(* Logix 5000 project; controller R400_500_XLS vendor 1 type 14 code 216 rev 31.11; software revision 31.01; part 12 of 32 *)
(* tags used below, declared in another part *)
   Chem_Pump : UDT_CHEM_PUMP[4];   // Chemical Pump flow rate
   CHEMICAL_COND_MAX_TIME : DINT;   // Timeout for the conductivity based chemical injection
   CHEMICAL_PUMP_OFF_TIME : DINT[4];
   CHEMICAL_PUMP_ON_TIME : DINT[4];
   FC87_CalibChemPmp : SINT;   // Calibration chemical pumps activation bits
   FC87_CalibChemPmpMsg : SINT;   // Chemical pump calibration step message
   FC87_ChemCalibRemainTime : DINT;
   FC87_ChemPumpIndex : SINT;   // Index of the selected chemical pump to calibrate
   FC87_LastValue : SINT;
   FC87_ONS : DINT;
   M : DINT[5];   // Memory Bits
   ONS_SPV17 : SINT;
   SET_POINT_FRACTION : REAL[4];
   Supervisor : DINT;
   Tmr : TIMER[107];
   ChemicalName : STRING[9];   // Used by HMI
   ChemPumpSelector : UDT_SELECTOR[2];   // Chemical pump calibration selector
   Current_Screen : DINT;
   DateTime : DINT[7];
   DateTimeNew : DINT[7];
   NumInput : UDT_NUMERIC_INPUT[65];   // Numeric input
   NumInputReal : UDT_NUMERIC_INPUT_REAL[17];
   RemoteDayOfMonth : DINT;   // HMI Date Day
   RemoteHour : DINT;   // HMI Time Hour
   RemoteMinute : DINT;   // HMI Time Minute
   RemoteMonth : DINT;   // HMI Date Month
   RemoteSecond : DINT;   // HMI Time Second
   RemoteSetDateTime : BOOL;   // HMI Set Date and Time
   RemoteYear : DINT;   // HMI Date Year
   Screen_Ctrl : DINT;   // PLC Screen Request
   SelChemi_Remote : SINT;
   SelChemical_Ind : SINT;
   SelChemical_Value : SINT;
   Selector : UDT_SELECTOR[25];   // Piloted list selector
   StringInput : UDT_STRING_INPUT[6];
   Tpb : DINT[11];
   TpbImage : DINT[11];
   Unit : Hrdwre;   // Unit Configuration
(* MainProgram, continued *)

ROUTINE SPV_12_CHEM_PUMP_CALIBRATION   (* ladder *)
// Calculate chemical pumps flow rate
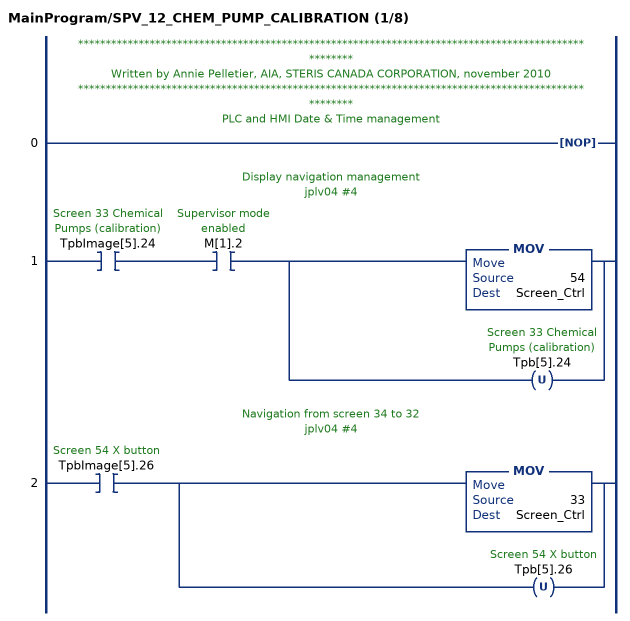
   // ****************************************************************************************************
   // Written by Annie Pelletier, AIA, STERIS CANADA CORPORATION, november 2010
   // ****************************************************************************************************
   // PLC and HMI Date & Time management
   0: NOP();
   // Display navigation management
   // jplv04 #4
   1: XIC(TpbImage[5].24)XIC(M[1].2)[MOV(54,Screen_Ctrl) ,OTU(Tpb[5].24) ];
   // Navigation from screen 34 to 32
   // jplv04 #4
   2: XIC(TpbImage[5].26)[MOV(33,Screen_Ctrl) ,OTU(Tpb[5].26) ];
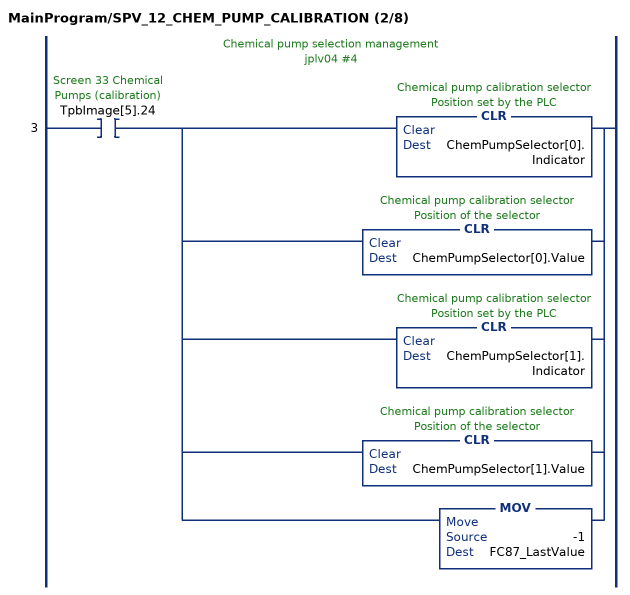
   // Chemical pump selection management
   // jplv04 #4
   3: XIC(TpbImage[5].24)[CLR(ChemPumpSelector[0].Indicator) ,CLR(ChemPumpSelector[0].Value) ,CLR(ChemPumpSelector[1].Indicator) ,CLR(ChemPumpSelector[1].Value) ,MOV(-1,FC87_LastValue) ];
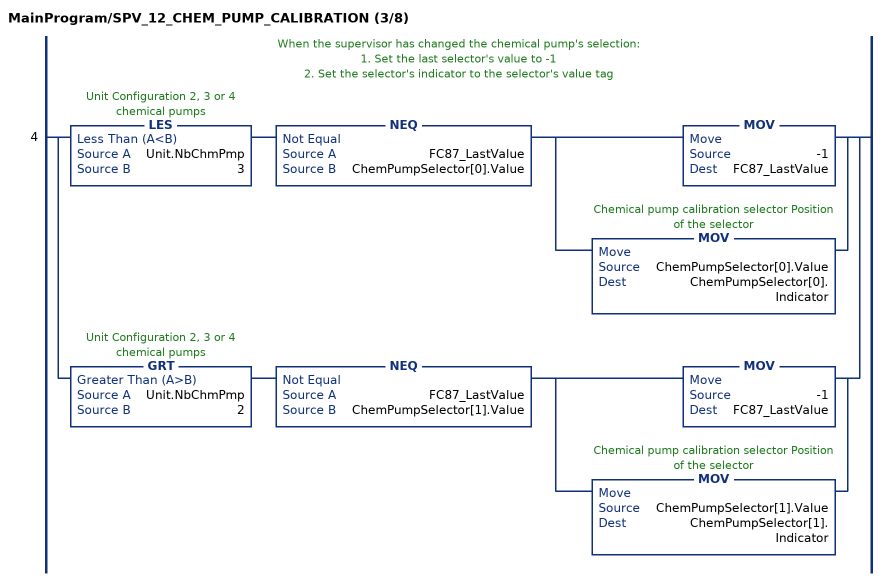
   // When the supervisor has changed the chemical pump's selection:
   // 1. Set the last selector's value to -1
   // 2. Set the selector's indicator to the selector's value tag
   4: [LES(Unit.NbChmPmp,3) NEQ(FC87_LastValue,ChemPumpSelector[0].Value) [MOV(-1,FC87_LastValue) ,MOV(ChemPumpSelector[0].Value,ChemPumpSelector[0].Indicator) ] ,GRT(Unit.NbChmPmp,2) NEQ(FC87_LastValue,ChemPumpSelector[1].Value) [MOV(-1,FC87_LastValue) ,MOV(ChemPumpSelector[1].Value,ChemPumpSelector[1].Indicator) ] ];
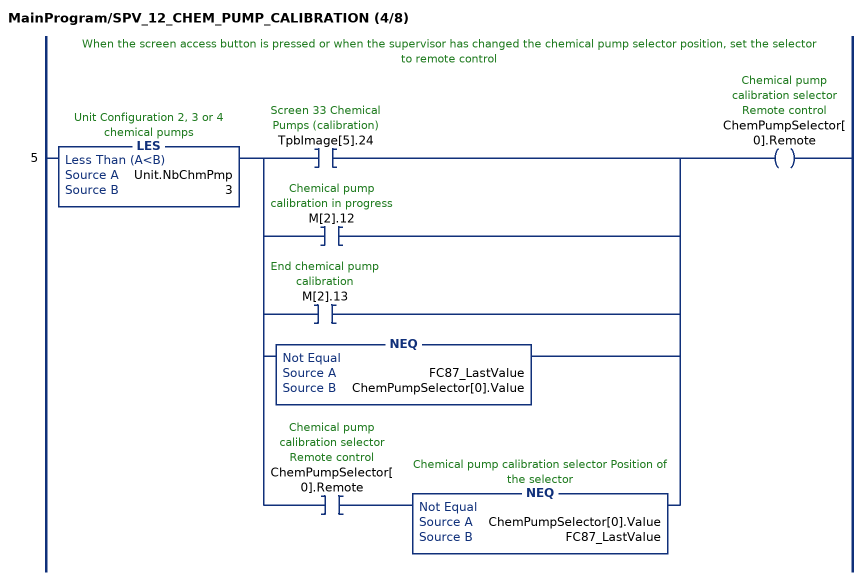
   // When the screen access button is pressed or when the supervisor has changed the chemical pump selector position, set the selector to remote control
   5: LES(Unit.NbChmPmp,3)[XIC(TpbImage[5].24) ,XIC(M[2].12) ,XIC(M[2].13) ,NEQ(FC87_LastValue,ChemPumpSelector[0].Value) ,XIC(ChemPumpSelector[0].Remote) NEQ(ChemPumpSelector[0].Value,FC87_LastValue) ]OTE(ChemPumpSelector[0].Remote);
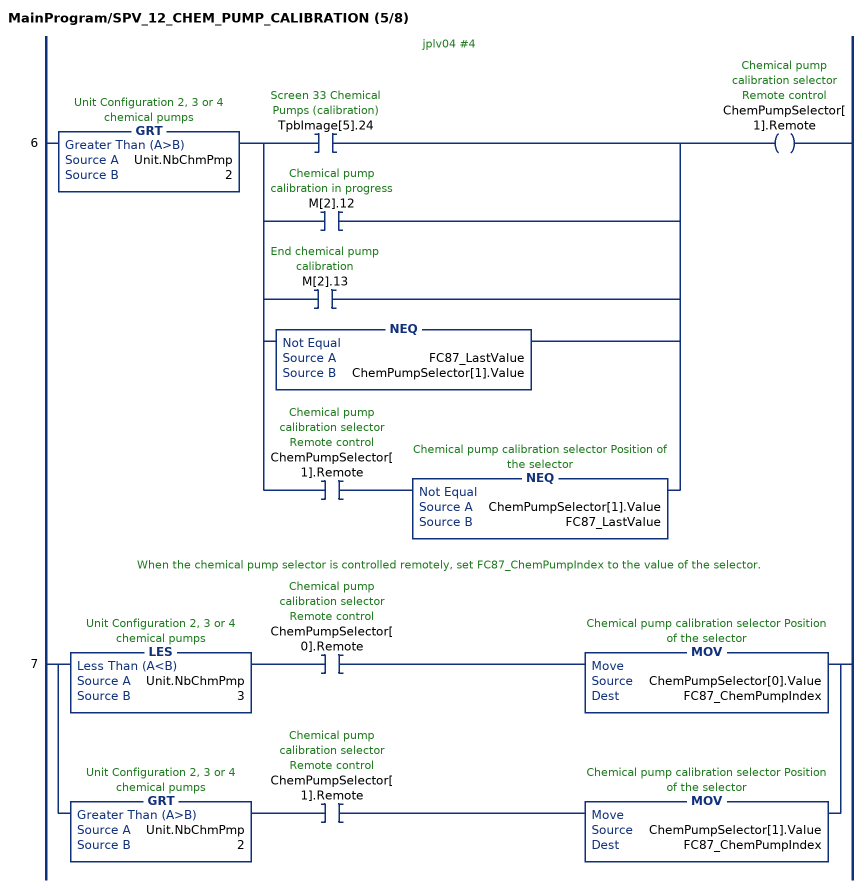
   // jplv04 #4
   6: GRT(Unit.NbChmPmp,2)[XIC(TpbImage[5].24) ,XIC(M[2].12) ,XIC(M[2].13) ,NEQ(FC87_LastValue,ChemPumpSelector[1].Value) ,XIC(ChemPumpSelector[1].Remote) NEQ(ChemPumpSelector[1].Value,FC87_LastValue) ]OTE(ChemPumpSelector[1].Remote);
   // When the chemical pump selector is controlled remotely, set FC87_ChemPumpIndex to the value of the selector.
   7: [LES(Unit.NbChmPmp,3) XIC(ChemPumpSelector[0].Remote) MOV(ChemPumpSelector[0].Value,FC87_ChemPumpIndex) ,GRT(Unit.NbChmPmp,2) XIC(ChemPumpSelector[1].Remote) MOV(ChemPumpSelector[1].Value,FC87_ChemPumpIndex) ];
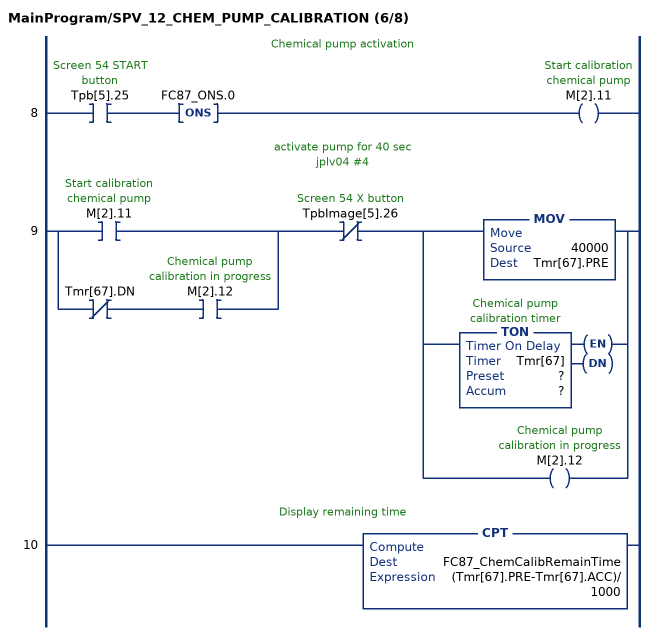
   // Chemical pump activation
   8: XIC(Tpb[5].25)ONS(FC87_ONS.0)OTE(M[2].11);
   // activate pump for 40 sec
   // jplv04 #4
   9: [XIC(M[2].11) ,XIO(Tmr[67].DN) XIC(M[2].12) ]XIO(TpbImage[5].26)[MOV(40000,Tmr[67].PRE) ,TON(Tmr[67],?,?) ,OTE(M[2].12) ];
   // Display remaining time
   10: CPT(FC87_ChemCalibRemainTime,(Tmr[67].PRE-Tmr[67].ACC)/1000);
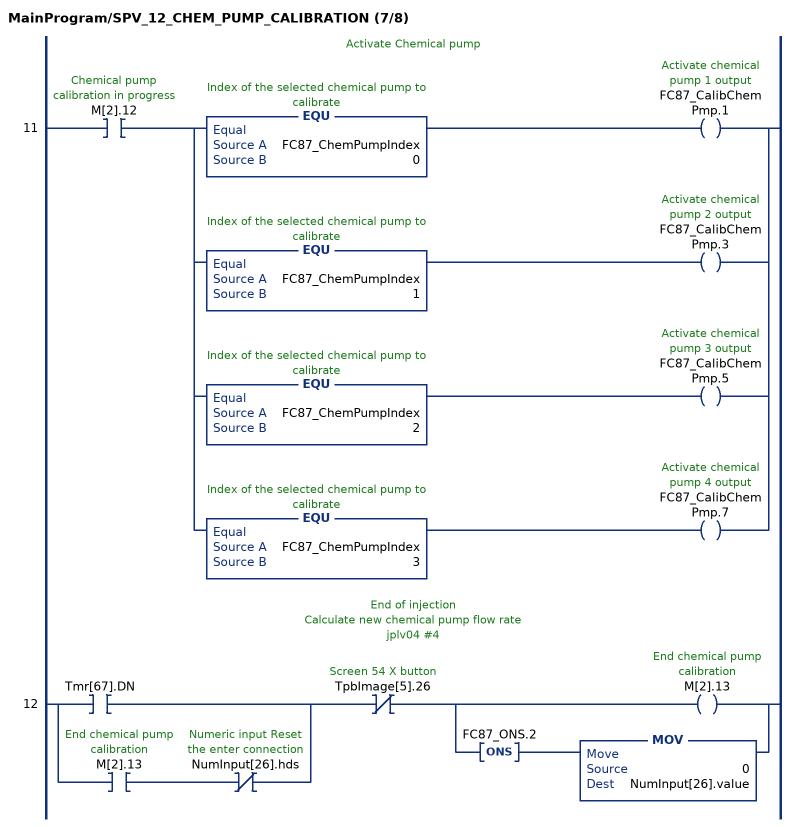
   // Activate Chemical pump
   11: XIC(M[2].12)[EQU(FC87_ChemPumpIndex,0) OTE(FC87_CalibChemPmp.1) ,EQU(FC87_ChemPumpIndex,1) OTE(FC87_CalibChemPmp.3) ,EQU(FC87_ChemPumpIndex,2) OTE(FC87_CalibChemPmp.5) ,EQU(FC87_ChemPumpIndex,3) OTE(FC87_CalibChemPmp.7) ];
   // End of injection
   // Calculate new chemical pump flow rate
   // jplv04 #4
   12: [XIC(Tmr[67].DN) ,XIC(M[2].13) XIO(NumInput[26].hds) ]XIO(TpbImage[5].26)[OTE(M[2].13) ,ONS(FC87_ONS.2) MOV(0,NumInput[26].value) ];
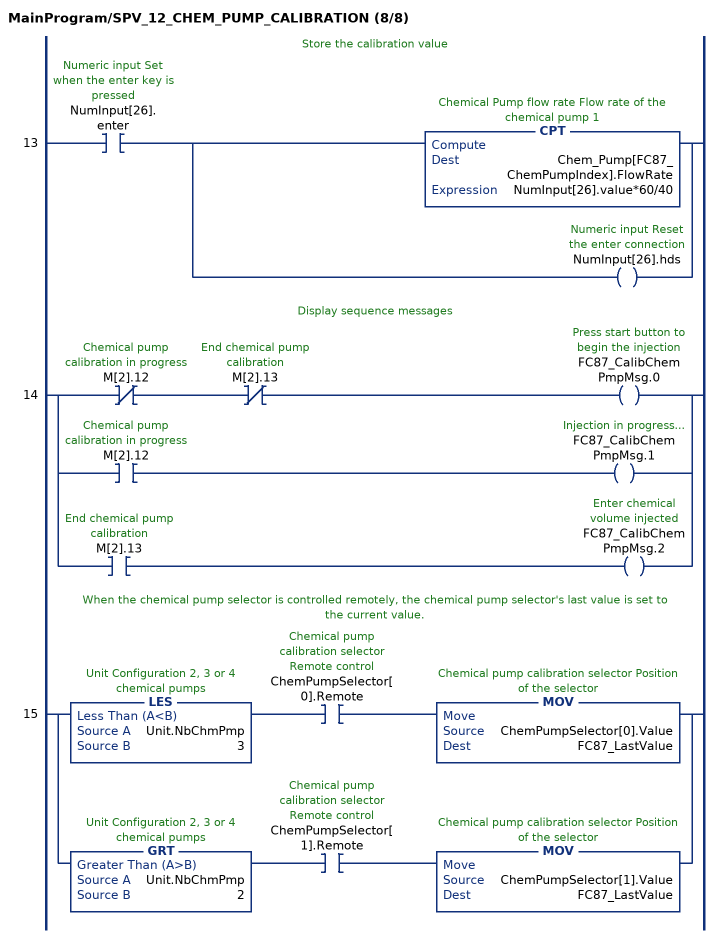
   // Store the calibration value
   13: XIC(NumInput[26].enter)[CPT(Chem_Pump[FC87_ChemPumpIndex].FlowRate,NumInput[26].value*60/40) ,OTE(NumInput[26].hds) ];
   // Display sequence messages
   14: [XIO(M[2].12) XIO(M[2].13) OTE(FC87_CalibChemPmpMsg.0) ,XIC(M[2].12) OTE(FC87_CalibChemPmpMsg.1) ,XIC(M[2].13) OTE(FC87_CalibChemPmpMsg.2) ];
   // When the chemical pump selector is controlled remotely, the chemical pump selector's last value is set to the current value.
   15: [LES(Unit.NbChmPmp,3) XIC(ChemPumpSelector[0].Remote) MOV(ChemPumpSelector[0].Value,FC87_LastValue) ,GRT(Unit.NbChmPmp,2) XIC(ChemPumpSelector[1].Remote) MOV(ChemPumpSelector[1].Value,FC87_LastValue) ];
END_ROUTINE

ROUTINE SPV_16_DATE_TIME   (* ladder *)
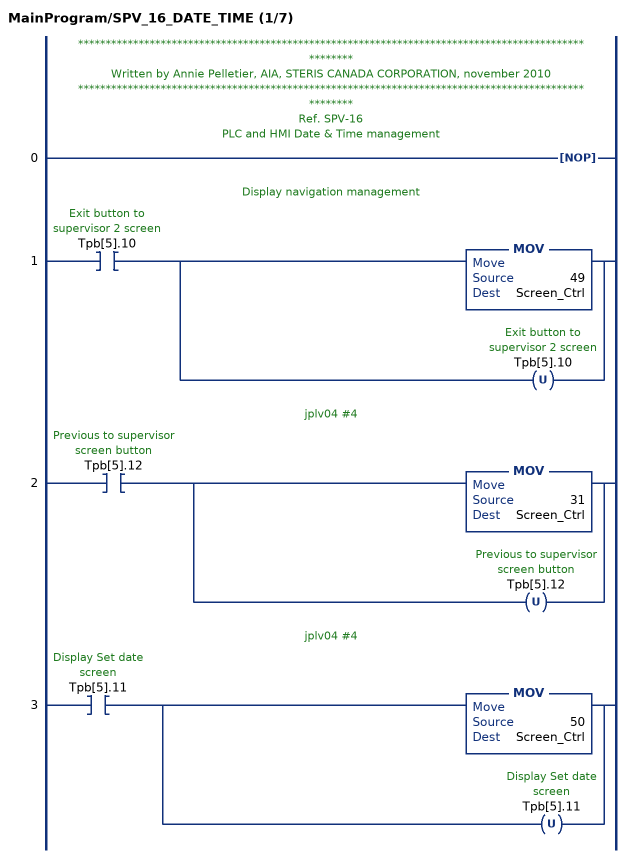
   // ****************************************************************************************************
   // Written by Annie Pelletier, AIA, STERIS CANADA CORPORATION, november 2010
   // ****************************************************************************************************
   // Ref. SPV-16
   // PLC and HMI Date & Time management
   0: NOP();
   // Display navigation management
   1: XIC(Tpb[5].10)[MOV(49,Screen_Ctrl) ,OTU(Tpb[5].10) ];
   // jplv04 #4
   2: XIC(Tpb[5].12)[MOV(31,Screen_Ctrl) ,OTU(Tpb[5].12) ];
   // jplv04 #4
   3: XIC(Tpb[5].11)[MOV(50,Screen_Ctrl) ,OTU(Tpb[5].11) ];
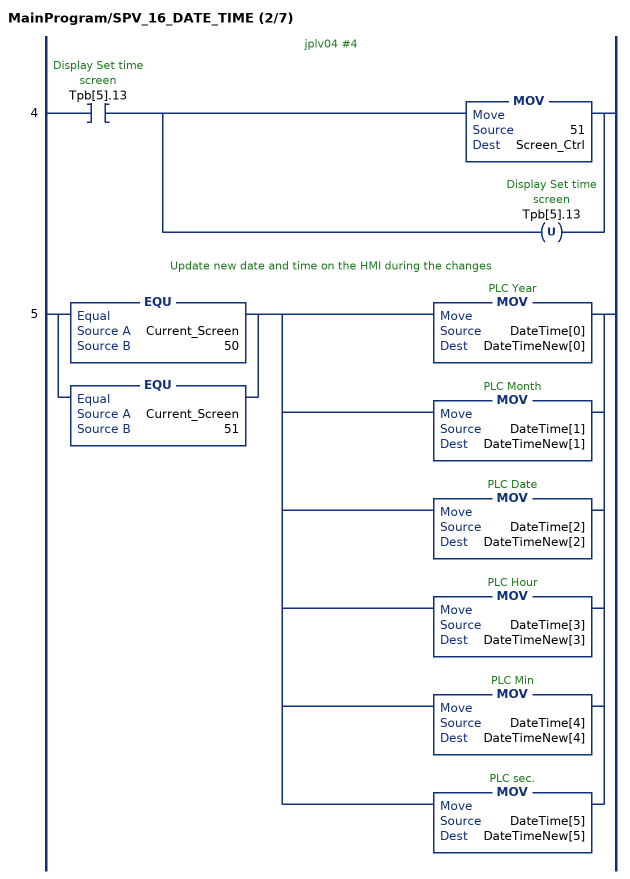
   // jplv04 #4
   4: XIC(Tpb[5].13)[MOV(51,Screen_Ctrl) ,OTU(Tpb[5].13) ];
   // Update new date and time on the HMI during the changes
   5: [EQU(Current_Screen,50) ,EQU(Current_Screen,51) ][MOV(DateTime[0],DateTimeNew[0]) ,MOV(DateTime[1],DateTimeNew[1]) ,MOV(DateTime[2],DateTimeNew[2]) ,MOV(DateTime[3],DateTimeNew[3]) ,MOV(DateTime[4],DateTimeNew[4]) ,MOV(DateTime[5],DateTimeNew[5]) ];
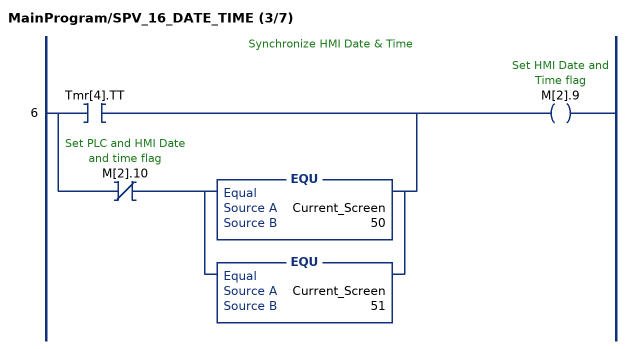
   // Synchronize HMI Date & Time
   6: [XIC(Tmr[4].TT) ,XIO(M[2].10) [EQU(Current_Screen,50) ,EQU(Current_Screen,51) ] ]OTE(M[2].9);
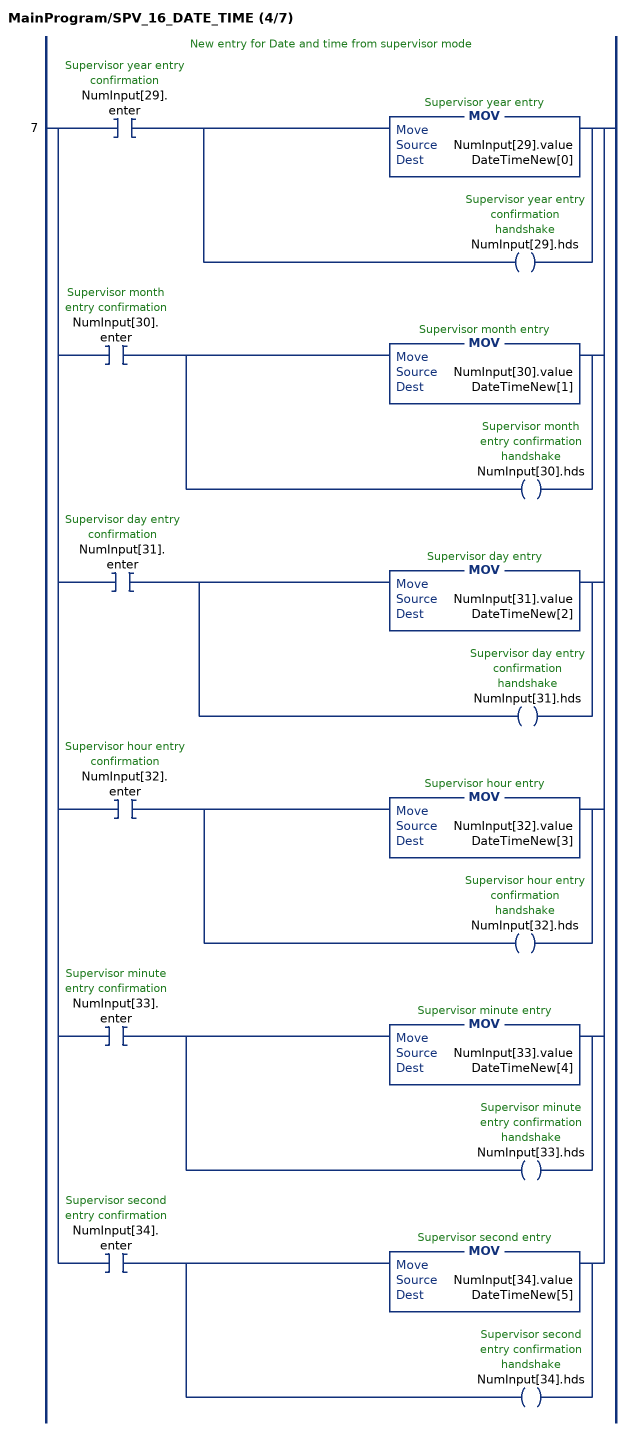
   // New entry for Date and time from supervisor mode
   7: [XIC(NumInput[29].enter) [MOV(NumInput[29].value,DateTimeNew[0]) ,OTE(NumInput[29].hds) ] ,XIC(NumInput[30].enter) [MOV(NumInput[30].value,DateTimeNew[1]) ,OTE(NumInput[30].hds) ] ,XIC(NumInput[31].enter) [MOV(NumInput[31].value,DateTimeNew[2]) ,OTE(NumInput[31].hds) ] ,XIC(NumInput[32].enter) [MOV(NumInput[32].value,DateTimeNew[3]) ,OTE(NumInput[32].hds) ] ,XIC(NumInput[33].enter) [MOV(NumInput[33].value,DateTimeNew[4]) ,OTE(NumInput[33].hds) ] ,XIC(NumInput[34].enter) [MOV(NumInput[34].value,DateTimeNew[5]) ,OTE(NumInput[34].hds) ] ];
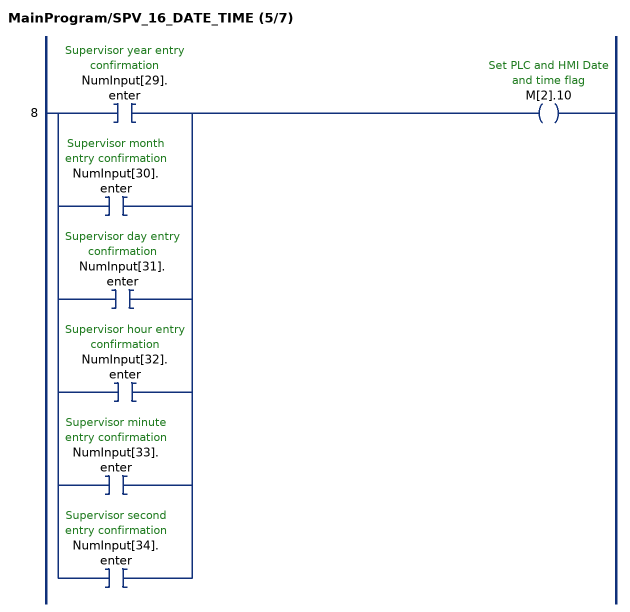
   8: [XIC(NumInput[29].enter) ,XIC(NumInput[30].enter) ,XIC(NumInput[31].enter) ,XIC(NumInput[32].enter) ,XIC(NumInput[33].enter) ,XIC(NumInput[34].enter) ]OTE(M[2].10);
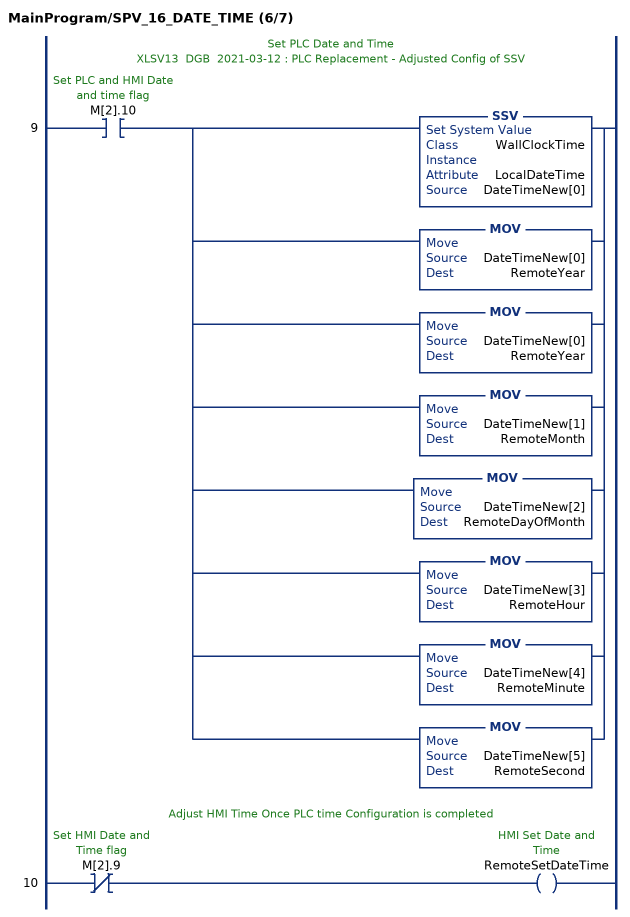
   // Set PLC Date and Time
   // XLSV13  DGB  2021-03-12 : PLC Replacement - Adjusted Config of SSV
   9: XIC(M[2].10)[SSV(WallClockTime,,LocalDateTime,DateTimeNew[0]) ,MOV(DateTimeNew[0],RemoteYear) ,MOV(DateTimeNew[0],RemoteYear) ,MOV(DateTimeNew[1],RemoteMonth) ,MOV(DateTimeNew[2],RemoteDayOfMonth) ,MOV(DateTimeNew[3],RemoteHour) ,MOV(DateTimeNew[4],RemoteMinute) ,MOV(DateTimeNew[5],RemoteSecond) ];
   // Adjust HMI Time Once PLC time Configuration is completed
   10: XIO(M[2].9)OTE(RemoteSetDateTime);
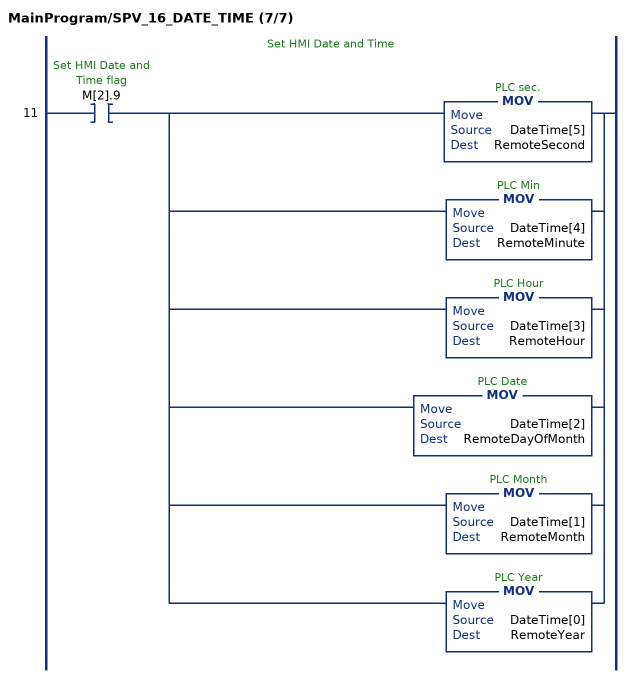
   // Set HMI Date and Time
   11: XIC(M[2].9)[MOV(DateTime[5],RemoteSecond) ,MOV(DateTime[4],RemoteMinute) ,MOV(DateTime[3],RemoteHour) ,MOV(DateTime[2],RemoteDayOfMonth) ,MOV(DateTime[1],RemoteMonth) ,MOV(DateTime[0],RemoteYear) ];
END_ROUTINE

ROUTINE SPV_17_Chemical_Parameters   (* ladder *)
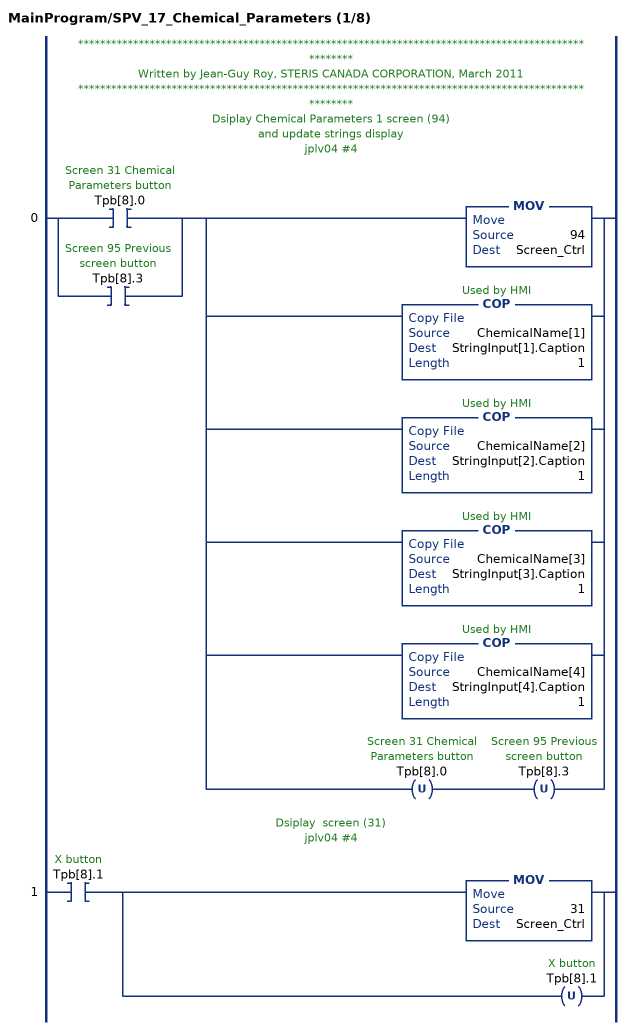
   // ****************************************************************************************************
   // Written by Jean-Guy Roy, STERIS CANADA CORPORATION, March 2011
   // ****************************************************************************************************
   // Dsiplay Chemical Parameters 1 screen (94)
   // and update strings display
   // jplv04 #4
   0: [XIC(Tpb[8].0) ,XIC(Tpb[8].3) ][MOV(94,Screen_Ctrl) ,COP(ChemicalName[1],StringInput[1].Caption,1) ,COP(ChemicalName[2],StringInput[2].Caption,1) ,COP(ChemicalName[3],StringInput[3].Caption,1) ,COP(ChemicalName[4],StringInput[4].Caption,1) ,OTU(Tpb[8].0) OTU(Tpb[8].3) ];
   // Dsiplay  screen (31)
   // jplv04 #4
   1: XIC(Tpb[8].1)[MOV(31,Screen_Ctrl) ,OTU(Tpb[8].1) ];
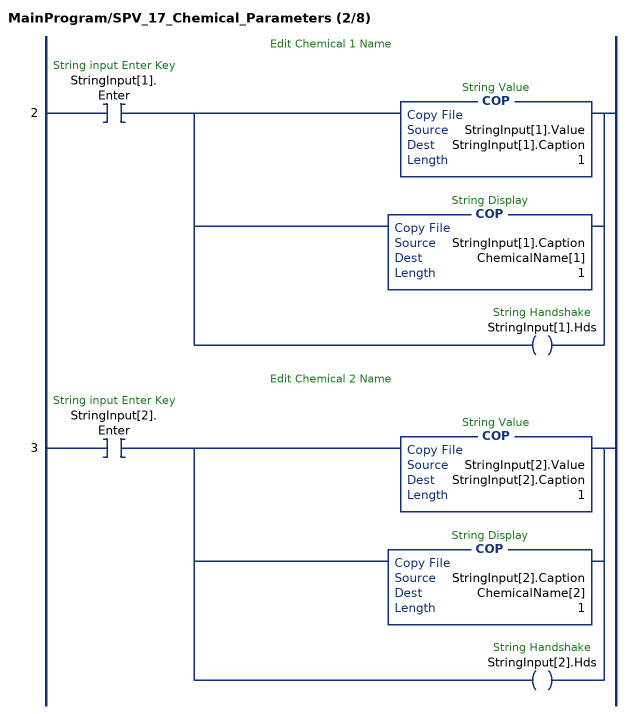
   // Edit Chemical 1 Name
   2: XIC(StringInput[1].Enter)[COP(StringInput[1].Value,StringInput[1].Caption,1) ,COP(StringInput[1].Caption,ChemicalName[1],1) ,OTE(StringInput[1].Hds) ];
   // Edit Chemical 2 Name
   3: XIC(StringInput[2].Enter)[COP(StringInput[2].Value,StringInput[2].Caption,1) ,COP(StringInput[2].Caption,ChemicalName[2],1) ,OTE(StringInput[2].Hds) ];
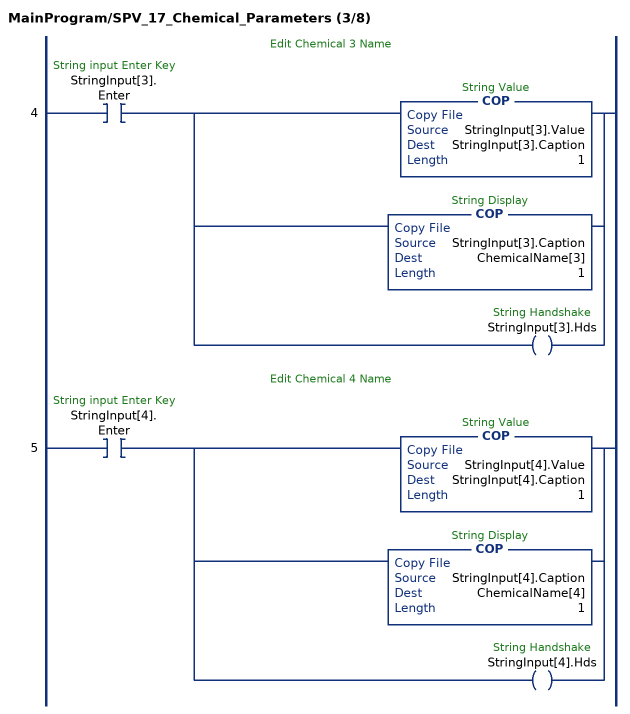
   // Edit Chemical 3 Name
   4: XIC(StringInput[3].Enter)[COP(StringInput[3].Value,StringInput[3].Caption,1) ,COP(StringInput[3].Caption,ChemicalName[3],1) ,OTE(StringInput[3].Hds) ];
   // Edit Chemical 4 Name
   5: XIC(StringInput[4].Enter)[COP(StringInput[4].Value,StringInput[4].Caption,1) ,COP(StringInput[4].Caption,ChemicalName[4],1) ,OTE(StringInput[4].Hds) ];
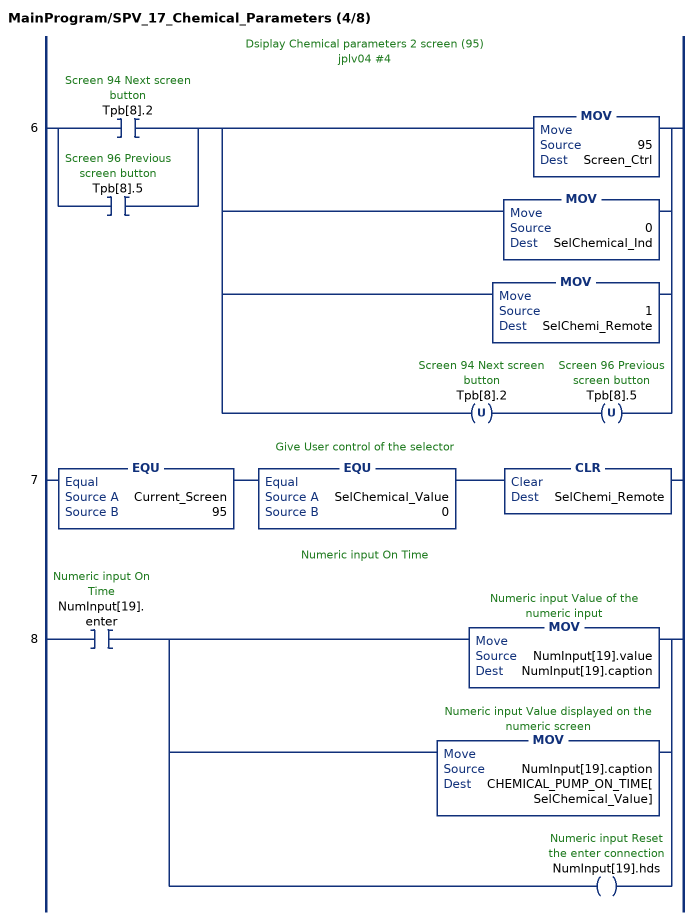
   // Dsiplay Chemical parameters 2 screen (95)
   // jplv04 #4
   6: [XIC(Tpb[8].2) ,XIC(Tpb[8].5) ][MOV(95,Screen_Ctrl) ,MOV(0,SelChemical_Ind) ,MOV(1,SelChemi_Remote) ,OTU(Tpb[8].2) OTU(Tpb[8].5) ];
   // Give User control of the selector
   7: EQU(Current_Screen,95)EQU(SelChemical_Value,0)CLR(SelChemi_Remote);
   // Numeric input On Time
   8: XIC(NumInput[19].enter)[MOV(NumInput[19].value,NumInput[19].caption) ,MOV(NumInput[19].caption,CHEMICAL_PUMP_ON_TIME[SelChemical_Value]) ,OTE(NumInput[19].hds) ];
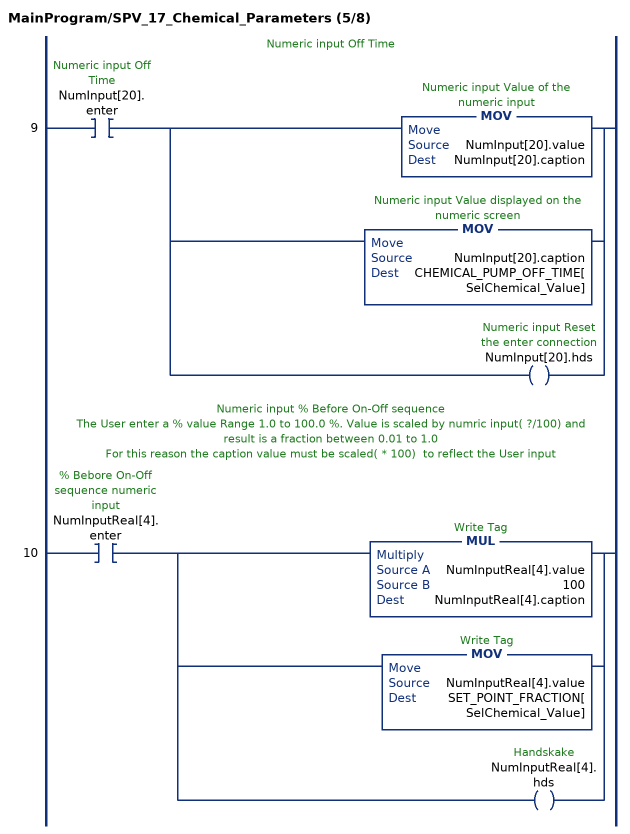
   // Numeric input Off Time
   9: XIC(NumInput[20].enter)[MOV(NumInput[20].value,NumInput[20].caption) ,MOV(NumInput[20].caption,CHEMICAL_PUMP_OFF_TIME[SelChemical_Value]) ,OTE(NumInput[20].hds) ];
   // Numeric input % Before On-Off sequence
   // The User enter a % value Range 1.0 to 100.0 %. Value is scaled by numric input( ?/100) and result is a fraction between 0.01 to 1.0
   // For this reason the caption value must be scaled( * 100)  to reflect the User input
   10: XIC(NumInputReal[4].enter)[MUL(NumInputReal[4].value,100,NumInputReal[4].caption) ,MOV(NumInputReal[4].value,SET_POINT_FRACTION[SelChemical_Value]) ,OTE(NumInputReal[4].hds) ];
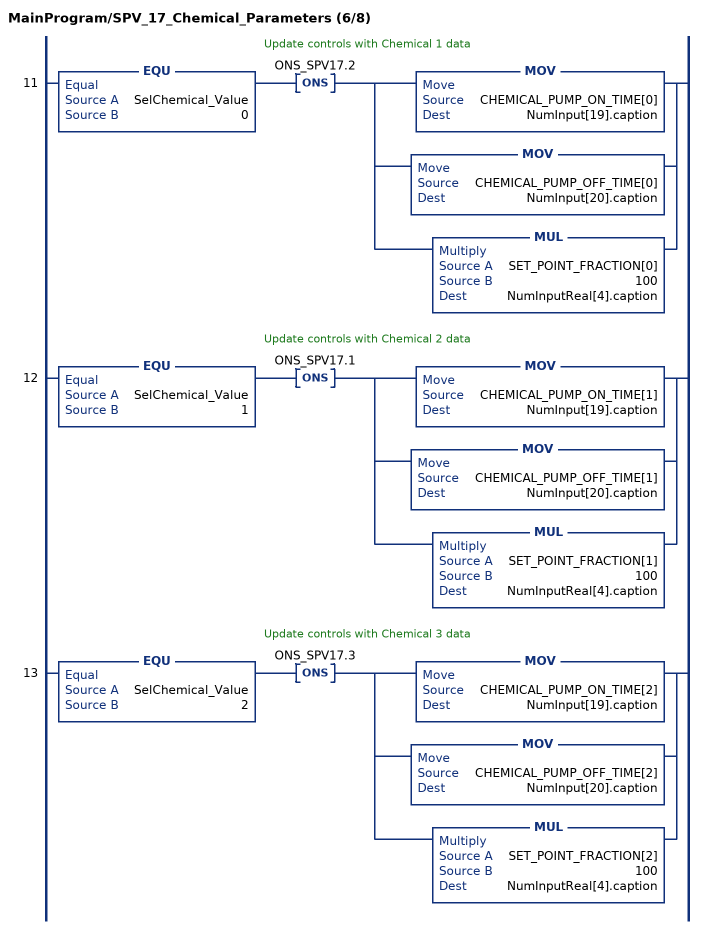
   // Update controls with Chemical 1 data
   11: EQU(SelChemical_Value,0)ONS(ONS_SPV17.2)[MOV(CHEMICAL_PUMP_ON_TIME[0],NumInput[19].caption) ,MOV(CHEMICAL_PUMP_OFF_TIME[0],NumInput[20].caption) ,MUL(SET_POINT_FRACTION[0],100,NumInputReal[4].caption) ];
   // Update controls with Chemical 2 data
   12: EQU(SelChemical_Value,1)ONS(ONS_SPV17.1)[MOV(CHEMICAL_PUMP_ON_TIME[1],NumInput[19].caption) ,MOV(CHEMICAL_PUMP_OFF_TIME[1],NumInput[20].caption) ,MUL(SET_POINT_FRACTION[1],100,NumInputReal[4].caption) ];
   // Update controls with Chemical 3 data
   13: EQU(SelChemical_Value,2)ONS(ONS_SPV17.3)[MOV(CHEMICAL_PUMP_ON_TIME[2],NumInput[19].caption) ,MOV(CHEMICAL_PUMP_OFF_TIME[2],NumInput[20].caption) ,MUL(SET_POINT_FRACTION[2],100,NumInputReal[4].caption) ];
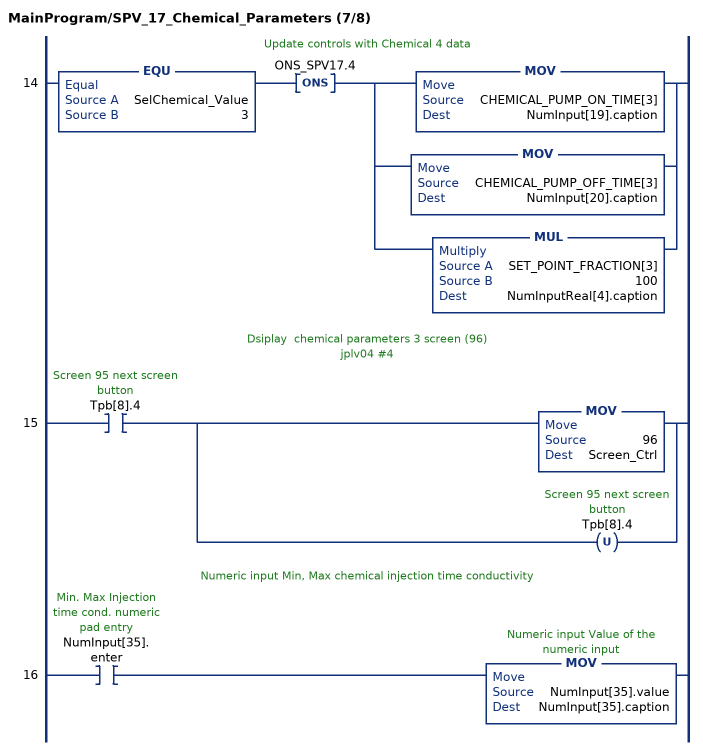
   // Update controls with Chemical 4 data
   14: EQU(SelChemical_Value,3)ONS(ONS_SPV17.4)[MOV(CHEMICAL_PUMP_ON_TIME[3],NumInput[19].caption) ,MOV(CHEMICAL_PUMP_OFF_TIME[3],NumInput[20].caption) ,MUL(SET_POINT_FRACTION[3],100,NumInputReal[4].caption) ];
   // Dsiplay  chemical parameters 3 screen (96)
   // jplv04 #4
   15: XIC(Tpb[8].4)[MOV(96,Screen_Ctrl) ,OTU(Tpb[8].4) ];
   // Numeric input Min, Max chemical injection time conductivity
   16: XIC(NumInput[35].enter)MOV(NumInput[35].value,NumInput[35].caption);
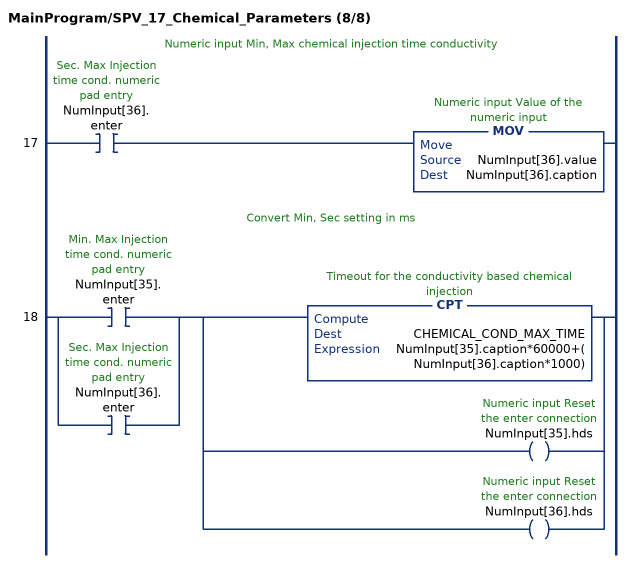
   // Numeric input Min, Max chemical injection time conductivity
   17: XIC(NumInput[36].enter)MOV(NumInput[36].value,NumInput[36].caption);
   // Convert Min, Sec setting in ms
   18: [XIC(NumInput[35].enter) ,XIC(NumInput[36].enter) ][CPT(CHEMICAL_COND_MAX_TIME,NumInput[35].caption*60000+(NumInput[36].caption*1000)) ,OTE(NumInput[35].hds) ,OTE(NumInput[36].hds) ];
END_ROUTINE
